(* IEC 61131-3 sources: Test-Git_ESME26/TestProgettoESME_26.fbsproj/AxisModuleLib Migration/DiagSource/AXM_FB_AxisModuleDiagSource.fb.st^ (part 2) *)

(* ---- WriteInterfaceMultiCamParamOut.meth.st ---- *)
METHOD INTERNAL WriteInterfaceMultiCamParamOut : BOOL
VAR_INPUT
END_VAR
VAR_OUTPUT
	q_etDiag		: GD.ET_Diag;
	q_etDiagExt	: TPL.ET_DiagExt;
	q_sMsg			: STRING[80];
END_VAR

THIS^.fbTreeWriter.Parameter(	i_sName		:= 'iq_xNewCam',
								i_sValue	:= BOOL_TO_STRING(THIS^.pstInterface^.stMultiCam.iq_xNewCam),
								q_etDiag	=> q_etDiag,
								q_etDiagExt	=> q_etDiagExt,
								q_sMsg		=> q_sMsg);

IF q_etDiag <> GD.ET_Diag.Ok THEN
	RETURN;
END_IF

THIS^.fbTreeWriter.Parameter(	i_sName		:= 'iq_xInstantNewCam',
								i_sValue	:= BOOL_TO_STRING(THIS^.pstInterface^.stMultiCam.iq_xInstantNewCam),
								q_etDiag	=> q_etDiag,
								q_etDiagExt	=> q_etDiagExt,
								q_sMsg		=> q_sMsg);

IF q_etDiag <> GD.ET_Diag.Ok THEN
	RETURN;
END_IF

THIS^.fbTreeWriter.Parameter(	i_sName		:= 'iq_xChangeMaster',
								i_sValue	:= BOOL_TO_STRING(THIS^.pstInterface^.stMultiCam.iq_xChangeMaster),
								q_etDiag	=> q_etDiag,
								q_etDiagExt	=> q_etDiagExt,
								q_sMsg		=> q_sMsg);

IF q_etDiag <> GD.ET_Diag.Ok THEN
	RETURN;
END_IF

THIS^.fbTreeWriter.Parameter(	i_sName		:= 'q_xXLowEnd',
								i_sValue	:= BOOL_TO_STRING(THIS^.pstInterface^.stMultiCam.q_xXLowEnd),
								q_etDiag	=> q_etDiag,
								q_etDiagExt	=> q_etDiagExt,
								q_sMsg		=> q_sMsg);

IF q_etDiag <> GD.ET_Diag.Ok THEN
	RETURN;
END_IF

THIS^.fbTreeWriter.Parameter(	i_sName		:= 'q_xXHighEnd',
								i_sValue	:= BOOL_TO_STRING(THIS^.pstInterface^.stMultiCam.q_xXHighEnd),
								q_etDiag	=> q_etDiag,
								q_etDiagExt	=> q_etDiagExt,
								q_sMsg		=> q_sMsg);

IF q_etDiag <> GD.ET_Diag.Ok THEN
	RETURN;
END_IF

THIS^.fbTreeWriter.Parameter(	i_sName		:= 'q_xInWsWindow',
								i_sValue	:= BOOL_TO_STRING(THIS^.pstInterface^.stMultiCam.q_xInWsWindow),
								q_etDiag	=> q_etDiag,
								q_etDiagExt	=> q_etDiagExt,
								q_sMsg		=> q_sMsg);

IF q_etDiag <> GD.ET_Diag.Ok THEN
	RETURN;
END_IF

THIS^.fbTreeWriter.Parameter(	i_sName		:= 'q_lrCalculatedCamPosition',
								i_sValue	:= LREAL_TO_STRING(THIS^.pstInterface^.stMultiCam.q_lrCalculatedCamPosition),
								q_etDiag	=> q_etDiag,
								q_etDiagExt	=> q_etDiagExt,
								q_sMsg		=> q_sMsg);

IF q_etDiag <> GD.ET_Diag.Ok THEN
	RETURN;
END_IF

THIS^.fbTreeWriter.Parameter(	i_sName		:= 'q_diActTable',
								i_sValue	:= DINT_TO_STRING(THIS^.pstInterface^.stMultiCam.q_diActTable),
								q_etDiag	=> q_etDiag,
								q_etDiagExt	=> q_etDiagExt,
								q_sMsg		=> q_sMsg);

IF q_etDiag <> GD.ET_Diag.Ok THEN
	RETURN;
END_IF

(* ---- WriteInterfaceMultiCamParamOutActualCamData.meth.st ---- *)
METHOD INTERNAL WriteInterfaceMultiCamParamOutActualCamData : BOOL
VAR_INPUT
END_VAR
VAR_OUTPUT
	q_etDiag		: GD.ET_Diag;
	q_etDiagExt	: TPL.ET_DiagExt;
	q_sMsg			: STRING[80];
END_VAR

THIS^.fbTreeWriter.NodeStart(	i_sName		:= 'q_stActualCamData',
								q_etDiag	=> q_etDiag,
								q_etDiagExt	=> q_etDiagExt,
								q_sMsg		=> q_sMsg);

IF q_etDiag <> GD.ET_Diag.Ok THEN
	RETURN;
END_IF

	THIS^.fbTreeWriter.Parameter(	i_sName		:= 'diProfileId',
									i_sValue	:= DINT_TO_STRING(THIS^.pstInterface^.stMultiCam.q_stActualCamData.diProfileId),
									q_etDiag	=> q_etDiag,
									q_etDiagExt	=> q_etDiagExt,
									q_sMsg		=> q_sMsg);

	IF q_etDiag <> GD.ET_Diag.Ok THEN
		RETURN;
	END_IF

	THIS^.fbTreeWriter.Parameter(	i_sName		:= 'lrXOffset',
									i_sValue	:= LREAL_TO_STRING(THIS^.pstInterface^.stMultiCam.q_stActualCamData.lrXOffset),
									q_etDiag	=> q_etDiag,
									q_etDiagExt	=> q_etDiagExt,
									q_sMsg		=> q_sMsg);

	IF q_etDiag <> GD.ET_Diag.Ok THEN
		RETURN;
	END_IF

	THIS^.fbTreeWriter.Parameter(	i_sName		:= 'lrYOffset',
									i_sValue	:= LREAL_TO_STRING(THIS^.pstInterface^.stMultiCam.q_stActualCamData.lrYOffset),
									q_etDiag	=> q_etDiag,
									q_etDiagExt	=> q_etDiagExt,
									q_sMsg		=> q_sMsg);

	IF q_etDiag <> GD.ET_Diag.Ok THEN
		RETURN;
	END_IF

	THIS^.fbTreeWriter.Parameter(	i_sName		:= 'lrXFactor',
									i_sValue	:= LREAL_TO_STRING(THIS^.pstInterface^.stMultiCam.q_stActualCamData.lrXFactor),
									q_etDiag	=> q_etDiag,
									q_etDiagExt	=> q_etDiagExt,
									q_sMsg		=> q_sMsg);

	IF q_etDiag <> GD.ET_Diag.Ok THEN
		RETURN;
	END_IF

	THIS^.fbTreeWriter.Parameter(	i_sName		:= 'lrYFactor',
									i_sValue	:= LREAL_TO_STRING(THIS^.pstInterface^.stMultiCam.q_stActualCamData.lrYFactor),
									q_etDiag	=> q_etDiag,
									q_etDiagExt	=> q_etDiagExt,
									q_sMsg		=> q_sMsg);

	IF q_etDiag <> GD.ET_Diag.Ok THEN
		RETURN;
	END_IF

	THIS^.fbTreeWriter.Parameter(	i_sName		:= 'diUserTableId',
									i_sValue	:= DINT_TO_STRING(THIS^.pstInterface^.stMultiCam.q_stActualCamData.diUserTableId),
									q_etDiag	=> q_etDiag,
									q_etDiagExt	=> q_etDiagExt,
									q_sMsg		=> q_sMsg);

	IF q_etDiag <> GD.ET_Diag.Ok THEN
		RETURN;
	END_IF

THIS^.fbTreeWriter.NodeEnd(	q_etDiag	=> q_etDiag,
							q_etDiagExt	=> q_etDiagExt,
							q_sMsg		=> q_sMsg);

IF q_etDiag <> GD.ET_Diag.Ok THEN
	RETURN;
END_IF

(* ---- WriteInterfaceMultiCamStart.meth.st ---- *)
METHOD INTERNAL WriteInterfaceMultiCamStart : BOOL
VAR_INPUT
END_VAR
VAR_OUTPUT
	q_etDiag		: GD.ET_Diag;
	q_etDiagExt	: TPL.ET_DiagExt;
	q_sMsg			: STRING[80];
END_VAR

THIS^.fbTreeWriter.NodeStart(	i_sName		:= 'stMultiCam',
								q_etDiag	=> q_etDiag,
								q_etDiagExt	=> q_etDiagExt,
								q_sMsg		=> q_sMsg);

(* ---- WriteInterfacePos.meth.st ---- *)
METHOD INTERNAL WriteInterfacePos : BOOL
VAR_INPUT
END_VAR
VAR_OUTPUT
	q_etDiag		: GD.ET_Diag;
	q_etDiagExt	: TPL.ET_DiagExt;
	q_sMsg			: STRING[80];
END_VAR

THIS^.fbTreeWriter.NodeStart(	i_sName		:= 'stPos',
								q_etDiag	=> q_etDiag,
								q_etDiagExt	=> q_etDiagExt,
								q_sMsg		=> q_sMsg);

IF q_etDiag <> GD.ET_Diag.Ok THEN
	RETURN;
END_IF

	THIS^.fbTreeWriter.Parameter(	i_sName		:= 'i_etPosMode',
									i_sValue	:= AXM_FC_EtPosModeToString(THIS^.pstInterface^.stPos.i_etPosMode),
									q_etDiag	=> q_etDiag,
									q_etDiagExt	=> q_etDiagExt,
									q_sMsg		=> q_sMsg);

	IF q_etDiag <> GD.ET_Diag.Ok THEN
		RETURN;
	END_IF

	THIS^.fbTreeWriter.Parameter(	i_sName		:= 'i_lrTarget',
									i_sValue	:= LREAL_TO_STRING(THIS^.pstInterface^.stPos.i_lrTarget),
									q_etDiag	=> q_etDiag,
									q_etDiagExt	=> q_etDiagExt,
									q_sMsg		=> q_sMsg);

	IF q_etDiag <> GD.ET_Diag.Ok THEN
		RETURN;
	END_IF

	THIS^.fbTreeWriter.Parameter(	i_sName		:= 'i_lrVel',
									i_sValue	:= LREAL_TO_STRING(THIS^.pstInterface^.stPos.i_lrVel),
									q_etDiag	=> q_etDiag,
									q_etDiagExt	=> q_etDiagExt,
									q_sMsg		=> q_sMsg);

	IF q_etDiag <> GD.ET_Diag.Ok THEN
		RETURN;
	END_IF

	THIS^.fbTreeWriter.Parameter(	i_sName		:= 'i_lrAcc',
									i_sValue	:= LREAL_TO_STRING(THIS^.pstInterface^.stPos.i_lrAcc),
									q_etDiag	=> q_etDiag,
									q_etDiagExt	=> q_etDiagExt,
									q_sMsg		=> q_sMsg);

	IF q_etDiag <> GD.ET_Diag.Ok THEN
		RETURN;
	END_IF

	THIS^.fbTreeWriter.Parameter(	i_sName		:= 'i_lrDec',
									i_sValue	:= LREAL_TO_STRING(THIS^.pstInterface^.stPos.i_lrDec),
									q_etDiag	=> q_etDiag,
									q_etDiagExt	=> q_etDiagExt,
									q_sMsg		=> q_sMsg);

	IF q_etDiag <> GD.ET_Diag.Ok THEN
		RETURN;
	END_IF

	THIS^.fbTreeWriter.Parameter(	i_sName		:= 'i_lrJerk',
									i_sValue	:= LREAL_TO_STRING(THIS^.pstInterface^.stPos.i_lrJerk),
									q_etDiag	=> q_etDiag,
									q_etDiagExt	=> q_etDiagExt,
									q_sMsg		=> q_sMsg);

	IF q_etDiag <> GD.ET_Diag.Ok THEN
		RETURN;
	END_IF

	THIS^.fbTreeWriter.Parameter(	i_sName		:= 'i_xStop',
									i_sValue	:= BOOL_TO_STRING(THIS^.pstInterface^.stPos.i_xStop),
									q_etDiag	=> q_etDiag,
									q_etDiagExt	=> q_etDiagExt,
									q_sMsg		=> q_sMsg);

	IF q_etDiag <> GD.ET_Diag.Ok THEN
		RETURN;
	END_IF

	THIS^.fbTreeWriter.Parameter(	i_sName		:= 'q_xInPosition',
									i_sValue	:= BOOL_TO_STRING(THIS^.pstInterface^.stPos.q_xInPosition),
									q_etDiag	=> q_etDiag,
									q_etDiagExt	=> q_etDiagExt,
									q_sMsg		=> q_sMsg);

	IF q_etDiag <> GD.ET_Diag.Ok THEN
		RETURN;
	END_IF

THIS^.fbTreeWriter.NodeEnd(	q_etDiag	=> q_etDiag,
							q_etDiagExt	=> q_etDiagExt,
							q_sMsg		=> q_sMsg);

IF q_etDiag <> GD.ET_Diag.Ok THEN
	RETURN;
END_IF

(* ---- WriteInterfaceStart.meth.st ---- *)
METHOD INTERNAL WriteInterfaceStart : BOOL
VAR_INPUT
END_VAR
VAR_OUTPUT
	q_etDiag		: GD.ET_Diag;
	q_etDiagExt	: TPL.ET_DiagExt;
	q_sMsg			: STRING[80];
END_VAR

THIS^.fbTreeWriter.NodeStart(	i_sName		:= 'ModuleInterface',
								q_etDiag	=> q_etDiag,
								q_etDiagExt	=> q_etDiagExt,
								q_sMsg		=> q_sMsg);
